(* IEC 61131-3 sources: llm-plc-st-eval/data/processed/gpt-4o/I1/zero_shot, 3 files *)

(* ---- ejec_1.st ---- *)
FUNCTION_BLOCK FB_Semaforo
VAR_INPUT
    habilitado : BOOL; // Entrada para habilitar o deshabilitar el semáforo
END_VAR_INPUT

VAR_OUTPUT
    luzV : BOOL; // Salida para la luz verde
    luzA : BOOL; // Salida para la luz amarilla
    luzR : BOOL; // Salida para la luz roja
END_VAR_OUTPUT

VAR
    estado : INT := 0; // Estado actual del semáforo
    temporizador : TON; // Temporizador para controlar los tiempos de cada luz
    parpadeo : BOOL := FALSE; // Estado del parpadeo amarillo
END_VAR

// Inicialización del temporizador
temporizador(IN := FALSE, PT := T#0S);

IF habilitado THEN
    // Secuencia cíclica del semáforo
    CASE estado OF
        0: // Luz verde
            luzV := TRUE;
            luzA := FALSE;
            luzR := FALSE;
            temporizador(IN := TRUE, PT := T#20S);
            IF temporizador.Q THEN
                estado := 1;
                temporizador(IN := FALSE);
            END_IF;
        1: // Luz amarilla
            luzV := FALSE;
            luzA := TRUE;
            luzR := FALSE;
            temporizador(IN := TRUE, PT := T#4S);
            IF temporizador.Q THEN
                estado := 2;
                temporizador(IN := FALSE);
            END_IF;
        2: // Luz roja
            luzV := FALSE;
            luzA := FALSE;
            luzR := TRUE;
            temporizador(IN := TRUE, PT := T#15S);
            IF temporizador.Q THEN
                estado := 0;
                temporizador(IN := FALSE);
            END_IF;
    END_CASE;
ELSE
    // Modo amarillo intermitente
    luzV := FALSE;
    luzR := FALSE;
    temporizador(IN := TRUE, PT := T#1S);
    IF temporizador.Q THEN
        parpadeo := NOT parpadeo;
        temporizador(IN := FALSE);
    END_IF;
    luzA := parpadeo;
    estado := 0; // Reiniciar la secuencia al habilitarse de nuevo
END_IF;
END_FUNCTION_BLOCK

(* ---- ejec_2.st ---- *)
FUNCTION_BLOCK FB_Semaforo
VAR_INPUT
    habilitado : BOOL; // Entrada para habilitar o deshabilitar el semáforo
END_VAR

VAR_OUTPUT
    luzV : BOOL; // Salida para la luz verde
    luzA : BOOL; // Salida para la luz amarilla
    luzR : BOOL; // Salida para la luz roja
END_VAR

VAR
    timer : TON; // Temporizador para controlar los tiempos de las luces
    estado : INT; // Estado actual del semáforo
    parpadeo : BOOL; // Estado de parpadeo para la luz amarilla
END_VAR

// Inicialización de variables
IF NOT habilitado THEN
    // Si no está habilitado, activar el modo intermitente amarillo
    luzV := FALSE;
    luzR := FALSE;
    timer(IN := TRUE, PT := T#1S);

    IF timer.Q THEN
        parpadeo := NOT parpadeo; // Alternar el estado de parpadeo
        timer(IN := FALSE); // Reiniciar el temporizador
    END_IF

    luzA := parpadeo; // Luz amarilla intermitente
    estado := 0; // Reiniciar el estado para cuando se habilite de nuevo
ELSE
    // Si está habilitado, seguir la secuencia normal del semáforo
    CASE estado OF
        0: // Estado de luz verde
            luzV := TRUE;
            luzA := FALSE;
            luzR := FALSE;
            timer(IN := TRUE, PT := T#20S);

            IF timer.Q THEN
                estado := 1; // Cambiar al estado de luz amarilla
                timer(IN := FALSE); // Reiniciar el temporizador
            END_IF

        1: // Estado de luz amarilla
            luzV := FALSE;
            luzA := TRUE;
            luzR := FALSE;
            timer(IN := TRUE, PT := T#4S);

            IF timer.Q THEN
                estado := 2; // Cambiar al estado de luz roja
                timer(IN := FALSE); // Reiniciar el temporizador
            END_IF

        2: // Estado de luz roja
            luzV := FALSE;
            luzA := FALSE;
            luzR := TRUE;
            timer(IN := TRUE, PT := T#15S);

            IF timer.Q THEN
                estado := 0; // Volver al estado de luz verde
                timer(IN := FALSE); // Reiniciar el temporizador
            END_IF
    END_CASE
END_IF
END_FUNCTION_BLOCK

(* ---- ejec_3.st ---- *)
FUNCTION_BLOCK FB_Semaforo
VAR
    // Variables de entrada
    habilitado : BOOL; // Indica si el semáforo está habilitado

    // Variables de salida
    luzV : BOOL := FALSE; // Luz verde
    luzA : BOOL := FALSE; // Luz amarilla
    luzR : BOOL := FALSE; // Luz roja

    // Variables internas
    estado : INT := 0; // Estado del semáforo
    temporizador : TON; // Temporizador para controlar los tiempos de las luces
    parpadeo : BOOL := FALSE; // Estado de parpadeo para luz amarilla intermitente
END_VAR

// Inicialización del temporizador
temporizador(IN := FALSE, PT := T#0S);

// Lógica del semáforo
IF habilitado THEN
    // Secuencia cíclica del semáforo
    CASE estado OF
        0: // Luz verde
            luzV := TRUE;
            luzA := FALSE;
            luzR := FALSE;
            temporizador(IN := TRUE, PT := T#20S);
            IF temporizador.Q THEN
                estado := 1;
                temporizador(IN := FALSE);
            END_IF;
        1: // Luz amarilla
            luzV := FALSE;
            luzA := TRUE;
            luzR := FALSE;
            temporizador(IN := TRUE, PT := T#4S);
            IF temporizador.Q THEN
                estado := 2;
                temporizador(IN := FALSE);
            END_IF;
        2: // Luz roja
            luzV := FALSE;
            luzA := FALSE;
            luzR := TRUE;
            temporizador(IN := TRUE, PT := T#15S);
            IF temporizador.Q THEN
                estado := 0;
                temporizador(IN := FALSE);
            END_IF;
    END_CASE;
ELSE
    // Luz amarilla intermitente
    luzV := FALSE;
    luzR := FALSE;
    temporizador(IN := TRUE, PT := T#1S);
    IF temporizador.Q THEN
        parpadeo := NOT parpadeo;
        temporizador(IN := FALSE);
    END_IF;
    luzA := parpadeo;
    estado := 0; // Reinicia el estado para comenzar en verde al habilitar
END_IF;
END_FUNCTION_BLOCK
